FUNCTION_BLOCK Algorithm_tu (* Basic Function Block Type *)
  (* Standard: 61499-2 *)
  (* Version 0.0, 10/23/2026, macie, Schneider Electric, Template *)
  PACKAGE Main;
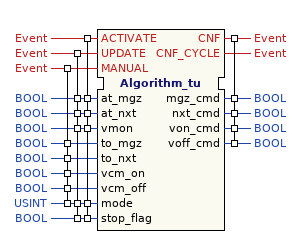
  EVENT_INPUT
    ACTIVATE WITH at_nxt, at_mgz, vmon, stop_flag, mode; (* Initialization Request *)
    UPDATE WITH at_nxt, at_mgz, vmon, stop_flag, mode; (* Normal Execution Request *)
    MANUAL WITH to_nxt, to_mgz, vcm_on, vcm_off, mode;
  END_EVENT
  EVENT_OUTPUT
    CNF WITH nxt_cmd, mgz_cmd, von_cmd, voff_cmd; (* Execution Confirmation *)
    CNF_CYCLE; (* Initialization Confirm *)
  END_EVENT
  VAR_INPUT
    at_mgz : BOOL;
    at_nxt : BOOL; (* Input event qualifier *)
    vmon : BOOL;
    to_mgz : BOOL;
    to_nxt : BOOL;
    vcm_on : BOOL;
    vcm_off : BOOL;
    mode : USINT;
    stop_flag : BOOL;
  END_VAR
  VAR_OUTPUT
    mgz_cmd : BOOL;
    nxt_cmd : BOOL; (* Output event qualifier *)
    von_cmd : BOOL;
    voff_cmd : BOOL;
  END_VAR
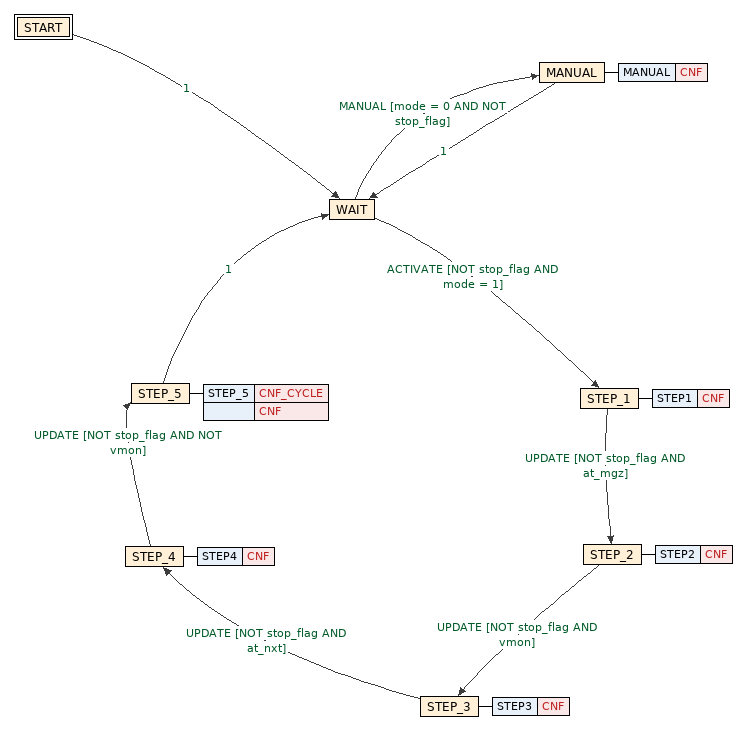
  EC_STATES
    START; (* Initial State *)
    WAIT;
    MANUAL : MANUAL -> CNF;
    STEP_1 : STEP1 -> CNF;
    STEP_2 : STEP2 -> CNF;
    STEP_3 : STEP3 -> CNF;
    STEP_4 : STEP4 -> CNF;
    STEP_5 : STEP_5 -> CNF_CYCLE, -> CNF;
  END_STATES
  EC_TRANSITIONS
    START TO WAIT := 1;
    WAIT TO MANUAL := MANUAL [mode = 0 AND NOT stop_flag];
    MANUAL TO WAIT := 1;
    WAIT TO STEP_1 := ACTIVATE [NOT stop_flag AND mode = 1];
    STEP_1 TO STEP_2 := UPDATE [NOT stop_flag AND at_mgz];
    STEP_2 TO STEP_3 := UPDATE [NOT stop_flag AND vmon];
    STEP_3 TO STEP_4 := UPDATE [NOT stop_flag AND at_nxt];
    STEP_4 TO STEP_5 := UPDATE [NOT stop_flag AND NOT vmon];
    STEP_5 TO WAIT := 1;
  END_TRANSITIONS
  ALGORITHM MANUAL IN ST:
;
nxt_cmd := to_nxt;
mgz_cmd := to_mgz;
von_cmd := vcm_on;
voff_cmd := vcm_off;
  END_ALGORITHM
  ALGORITHM STEP1 IN ST:
;
mgz_cmd := TRUE;
nxt_cmd := FALSE;
  END_ALGORITHM
  ALGORITHM STEP2 IN ST:
;
von_cmd := TRUE;
voff_cmd := FALSE;
  END_ALGORITHM
  ALGORITHM STEP3 IN ST:
;
nxt_cmd := TRUE;
mgz_cmd := FALSE;
  END_ALGORITHM
  ALGORITHM STEP4 IN ST:
;
voff_cmd := TRUE;
von_cmd := FALSE;
  END_ALGORITHM
  ALGORITHM STEP_5 IN ST:
;
vcm_off := FALSE;
  END_ALGORITHM
END_FUNCTION_BLOCK
